// TwinCAT 3 PLC project Untitled1
// ProgramVersion: 3.1.4024.0
// libraries:
//   Tc2_Standard, * (Beckhoff Automation GmbH)
//   Tc2_System, * (Beckhoff Automation GmbH)
//   Tc3_Module, * (Beckhoff Automation GmbH)
// project tree:
//   / PlcTask.TcTTO
//   POUs/ PLC_PRG.TcPOU, VltFixtureCfc.TcPOU, VltFixtureSfc.TcPOU
// real-time tasks:
//   TASK PlcTask: cycle T#10ms, priority 20, ADS port 350

CONFIGURATION Untitled1
    RESOURCE PLC ON TwinCAT3
        TASK PlcTask(INTERVAL := T#10ms, PRIORITY := 20);
        PROGRAM PLC_PRG WITH PlcTask : PLC_PRG;
    END_RESOURCE
END_CONFIGURATION

// ---- POUs/PLC_PRG.TcPOU
PROGRAM PLC_PRG
VAR


END_VAR

END_PROGRAM

// ---- POUs/VltFixtureCfc.TcPOU
PROGRAM VltFixtureCfc
VAR
END_VAR

END_PROGRAM

// ---- POUs/VltFixtureSfc.TcPOU
PROGRAM VltFixtureSfc
VAR
END_VAR

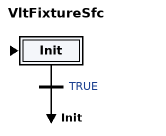
INITIAL_STEP Init:
END_STEP
TRANSITION FROM Init TO Init
    := TRUE;
END_TRANSITION

END_PROGRAM
